(* IEC 61131-3 sources: podajnik-arkuszy/plc, 8 files *)

(* ---- FB_EStop.st ---- *)
(* Zezwolenie ruchu. Po otwarciu obwodu bezpieczenstwa i po wlaczeniu zasilania
   wymagane jest zbocze kasowania. Sam powrot styku bezpieczenstwa nie uruchamia maszyny. *)
FUNCTION_BLOCK FB_EStop
VAR_INPUT
    EStopOk : BOOL;
    Reset : BOOL;
END_VAR
VAR_OUTPUT
    RunEnable : BOOL;
END_VAR
VAR
    NeedReset : BOOL := TRUE;
END_VAR

IF NOT EStopOk THEN
    NeedReset := TRUE;
    RunEnable := FALSE;
ELSIF NeedReset THEN
    RunEnable := FALSE;
    IF Reset THEN
        NeedReset := FALSE;
        RunEnable := TRUE;
    END_IF;
ELSE
    RunEnable := TRUE;
END_IF;

END_FUNCTION_BLOCK

(* ---- FB_FuserBuckle.st ---- *)
(* Predkosc silnika fusera od czujnika wybrzuszenia przed nipem.
   Za duze wybrzuszenie: przyspiesz, zeby nie zgniesc arkusza.
   Za male: zwolnij, zeby nie rozmazac toneru na pasie.
   Waskie medium obcina predkosc. Zawiniecie na pasie zatrzymuje naped. *)
FUNCTION_BLOCK FB_FuserBuckle
VAR_INPUT
    Enable : BOOL;
    Nip : BOOL;
    BuckleHigh : BOOL;
    BuckleLow : BOOL;
    NarrowMedia : BOOL;
    Wrap : BOOL;
END_VAR
VAR_OUTPUT
    SpeedPct : INT;
    HeaterOn : BOOL;
    Jam : BOOL;
END_VAR

IF NOT Enable OR Wrap THEN
    SpeedPct := 0;
    HeaterOn := FALSE;
    Jam := Wrap;
ELSE
    Jam := FALSE;
    HeaterOn := TRUE; (* ceramika w pasie *)
    SpeedPct := 100;

    IF Nip AND BuckleHigh THEN
        SpeedPct := 130;
    ELSIF Nip AND BuckleLow THEN
        SpeedPct := 70;
    END_IF;

    IF NarrowMedia AND (SpeedPct > 80) THEN
        SpeedPct := 80;
    END_IF;
END_IF;

END_FUNCTION_BLOCK

(* ---- FB_FuserLife.st ---- *)
(* Licznik fusera. W XC4140 komplet type 01 (41X0253) wymienia sie po 150 000 stron.
   Ostrzezenie od 140 000. Kasowanie jest osobne od resetu zaciecia.
   Na panel idzie liczba tysiecy: rejestr 16-bit nie zmiesci 150000. *)
FUNCTION_BLOCK FB_FuserLife
VAR_INPUT
    SheetCount : INT;
    ResetService : BOOL;
END_VAR
VAR_OUTPUT
    Thousands : INT;
    Warn : BOOL;
    Due : BOOL;
END_VAR
VAR
    Total : DINT := 0;
    Prev : INT := 0;
    Seen : BOOL := FALSE;
END_VAR

IF NOT Seen THEN
    Prev := SheetCount;
    Seen := TRUE;
END_IF;

IF ResetService THEN
    Total := 0;
ELSIF SheetCount <> Prev THEN
    Total := Total + 1;
END_IF;
Prev := SheetCount;

IF Total > 150000 THEN
    Total := 150000;
END_IF;

Thousands := DINT_TO_INT(Total / 1000);
Warn := Total >= 140000;
Due := Total >= 150000;

END_FUNCTION_BLOCK

(* ---- FB_Motor.st ---- *)
(* Stycznik silnika. FaultIn przychodzi z termika.
   Gdy UseFeedback = TRUE, brak styku pomocniczego dluzej niz 500 ms jest awaria napedu. *)
FUNCTION_BLOCK FB_Motor
VAR_INPUT
    RunCmd : BOOL;
    Feedback : BOOL;
    UseFeedback : BOOL;
    FaultIn : BOOL;
    Reset : BOOL;
END_VAR
VAR_OUTPUT
    Run : BOOL;
    Fault : BOOL;
END_VAR
VAR
    TonFb : TON;
END_VAR

IF FaultIn THEN
    Fault := TRUE;
END_IF;

IF Reset AND NOT FaultIn THEN
    Fault := FALSE;
END_IF;

IF Fault THEN
    Run := FALSE;
    TonFb(IN := FALSE, PT := T#500ms);
ELSE
    IF UseFeedback THEN
        TonFb(IN := RunCmd AND NOT Feedback, PT := T#500ms);
    ELSE
        TonFb(IN := FALSE, PT := T#500ms);
    END_IF;

    IF TonFb.Q THEN
        Fault := TRUE;
        Run := FALSE;
    ELSE
        Run := RunCmd;
    END_IF;
END_IF;

END_FUNCTION_BLOCK

(* ---- FB_PID.st ---- *)
(* Regulator grzalki 24 V. Wyjscie 0..100 procent.
   Pierwszy cykl po wlaczeniu nie daje kopa od czlonu D. *)
FUNCTION_BLOCK FB_PID
VAR_INPUT
    Enable : BOOL;
    Setpoint : REAL;
    Actual : REAL;
    Kp : REAL;
    Ki : REAL;
    Kd : REAL;
    OutMin : REAL;
    OutMax : REAL;
    Cycle : REAL; (* okres obiegu w sekundach, przy cyklu 10 ms wpisz 0.01 *)
END_VAR
VAR_OUTPUT
    Out : REAL;
END_VAR
VAR
    Integral : REAL := 0.0;
    PrevError : REAL := 0.0;
    Armed : BOOL := FALSE;
    Error : REAL;
    Deriv : REAL;
    Raw : REAL;
END_VAR

IF NOT Enable OR (Cycle <= 0.0) THEN
    Integral := 0.0;
    PrevError := 0.0;
    Armed := FALSE;
    Out := 0.0;
ELSE
    Error := Setpoint - Actual;
    IF NOT Armed THEN
        PrevError := Error;
        Integral := 0.0;
        Armed := TRUE;
    END_IF;

    Integral := Integral + (Error * Cycle);
    Deriv := (Error - PrevError) / Cycle;
    PrevError := Error;
    Raw := (Kp * Error) + (Ki * Integral) + (Kd * Deriv);

    IF Raw > OutMax THEN
        Raw := OutMax;
        Integral := Integral - (Error * Cycle);
    ELSIF Raw < OutMin THEN
        Raw := OutMin;
        Integral := Integral - (Error * Cycle);
    END_IF;

    Out := Raw;
END_IF;

END_FUNCTION_BLOCK

(* ---- FB_SheetTrack.st ---- *)
(* Sciezka arkusza: sprzeglo podaje, czujnik wejscia, rejestracja, czujnik wyjscia.
   Brak czujnika w czasie JamTime (domyslnie 800 ms) = zaciecie.
   Przerwanie cyklu, gdy arkusz jest jeszcze na czujniku, tez jest zacieciem.
   Kasowanie dziala tylko przy pustej sciezce. *)
FUNCTION_BLOCK FB_SheetTrack
VAR_INPUT
    FeedCmd : BOOL;
    SensEntry : BOOL;
    SensRegister : BOOL;
    SensExit : BOOL;
    Reset : BOOL;
    JamTime : TIME := T#800ms;
END_VAR
VAR_OUTPUT
    MotorCmd : BOOL;
    Clutch : BOOL;
    AtRegister : BOOL;
    Jam : BOOL;
    Busy : BOOL;
    SheetCount : INT;
    PhaseOut : INT;
END_VAR
VAR
    Phase : INT := 0; (* 0 postoj, 1 czekam na rejestracje, 2 przejazd, 3 zejscie z czujnika *)
    TonReg : TON;
    TonExit : TON;
    rEntry : R_TRIG;
    rExit : R_TRIG;
END_VAR

rEntry(CLK := SensEntry);
rExit(CLK := SensExit);
TonReg(IN := (Phase = 1) AND NOT Jam, PT := JamTime);
TonExit(IN := (Phase = 2) AND NOT Jam, PT := JamTime);

IF Reset AND NOT SensEntry AND NOT SensRegister AND NOT SensExit THEN
    Jam := FALSE;
    Phase := 0;
END_IF;

IF Jam THEN
    MotorCmd := FALSE;
    Clutch := FALSE;
    AtRegister := FALSE;
ELSIF NOT FeedCmd AND (Phase <> 0) THEN
    IF SensEntry OR SensRegister OR SensExit THEN
        Jam := TRUE;
    ELSE
        Phase := 0;
    END_IF;
    MotorCmd := FALSE;
    Clutch := FALSE;
    AtRegister := FALSE;
ELSIF Phase = 0 THEN
    AtRegister := FALSE;
    IF FeedCmd AND rEntry.Q THEN
        Clutch := FALSE;
        MotorCmd := TRUE;
        Phase := 1;
    ELSIF FeedCmd AND (SensEntry OR SensRegister OR SensExit) THEN
        Jam := TRUE;
        Clutch := FALSE;
        MotorCmd := FALSE;
    ELSIF FeedCmd THEN
        Clutch := TRUE;
        MotorCmd := TRUE;
    ELSE
        Clutch := FALSE;
        MotorCmd := FALSE;
    END_IF;
ELSIF Phase = 1 THEN
    Clutch := FALSE;
    MotorCmd := TRUE;
    AtRegister := FALSE;
    IF SensRegister THEN
        Phase := 2;
        AtRegister := TRUE;
    ELSIF TonReg.Q THEN
        Jam := TRUE;
        Phase := 0;
        MotorCmd := FALSE;
    END_IF;
ELSIF Phase = 2 THEN
    Clutch := FALSE;
    MotorCmd := TRUE;
    AtRegister := TRUE;
    IF rExit.Q THEN
        SheetCount := SheetCount + 1;
        Phase := 3;
        AtRegister := FALSE;
    ELSIF TonExit.Q THEN
        Jam := TRUE;
        Phase := 0;
        MotorCmd := FALSE;
        AtRegister := FALSE;
    END_IF;
ELSE
    Clutch := FALSE;
    AtRegister := FALSE;
    MotorCmd := TRUE;
    IF NOT SensExit AND NOT SensEntry AND NOT SensRegister THEN
        Phase := 0;
        MotorCmd := FALSE;
    END_IF;
END_IF;

IF Jam THEN
    MotorCmd := FALSE;
    Clutch := FALSE;
    AtRegister := FALSE;
END_IF;

Busy := Jam OR (Phase <> 0) OR Clutch;
PhaseOut := Phase;

END_FUNCTION_BLOCK

(* ---- FB_Warmup.st ---- *)
(* Zezwolenie na podanie, gdy rolka 24 V jest w pasmie.
   Zadanie regulatora to 80 C. Ponizej 70 C start jest martwy.
   Powyzej 95 C to przegrzanie: grzalka odpada, nowy arkusz tez. *)
FUNCTION_BLOCK FB_Warmup
VAR_INPUT
    Enable : BOOL;
    Actual : REAL;
END_VAR
VAR_OUTPUT
    Ready : BOOL;
    Heating : BOOL;
    Overtemp : BOOL;
END_VAR

Overtemp := Enable AND (Actual > 95.0);
Ready := Enable AND (Actual >= 70.0) AND (Actual <= 95.0);
Heating := Enable AND (Actual < 70.0);

END_FUNCTION_BLOCK

(* ---- MAIN.st ---- *)
(* Podajnik arkuszy.
   OpenPLC Editor albo CODESYS: wklej FB_*.st jako bloki funkcyjne, a ten plik jako program.
   Cykl zadania: 10 ms.
   Adresy sa zgodne z electrical/io_map.csv.
   UseFeedback ustaw na TRUE dopiero po podpieciu styku pomocniczego stycznika pod I_MotorAux. *)
PROGRAM Main
VAR
    I_EstopOk AT %IX0.0 : BOOL;
    I_CoverClosed AT %IX0.1 : BOOL;
    I_SensEntry AT %IX0.2 : BOOL;
    I_SensRegister AT %IX0.3 : BOOL;
    I_SensExit AT %IX0.4 : BOOL;
    I_MotorFault AT %IX0.5 : BOOL;
    I_Start AT %IX0.6 : BOOL;
    I_Stop AT %IX0.7 : BOOL;
    I_Reset AT %IX1.0 : BOOL;
    I_MotorAux AT %IX1.1 : BOOL;
    I_FuserReset AT %IX1.2 : BOOL;
    I_Nip AT %IX1.3 : BOOL;
    I_BuckleHigh AT %IX1.4 : BOOL;
    I_BuckleLow AT %IX1.5 : BOOL;
    I_NarrowMedia AT %IX1.6 : BOOL;
    I_FuserWrap AT %IX1.7 : BOOL;
    IW_TempRaw AT %IW2 : INT;

    Q_Motor AT %QX0.0 : BOOL;
    Q_Clutch AT %QX0.1 : BOOL;
    Q_Gate AT %QX0.2 : BOOL;
    Q_LampRun AT %QX0.3 : BOOL;
    Q_LampFault AT %QX0.4 : BOOL;
    Q_Heater AT %QX0.5 : BOOL;
    Q_FuserMotor AT %QX0.6 : BOOL;

    QW_Heater AT %QW0 : INT; (* 0..1000 = 0.0..100.0 % *)
    QW_State AT %QW1 : INT;
    QW_Sheets AT %QW2 : INT;
    QW_Temp AT %QW3 : INT;
    QW_FuserK AT %QW4 : INT; (* tysiace stron od resetu fusera *)
    QW_FuserSvc AT %QW5 : INT; (* 0 ok, 1 ostrzezenie, 2 wymiana *)
    QW_FuserSpeed AT %QW6 : INT; (* procent predkosci silnika fusera *)
    QW_Warm AT %QW7 : INT; (* 0 zimna, 1 gotowa, 2 przegrzanie *)

    EStop : FB_EStop;
    Drive : FB_Motor;
    Track : FB_SheetTrack;
    Heat : FB_PID;
    FuserLife : FB_FuserLife;
    Buckle : FB_FuserBuckle;
    Warmup : FB_Warmup;
    rStart : R_TRIG;
    rStop : R_TRIG;
    rReset : R_TRIG;
    RunRequest : BOOL := FALSE;
    UseFeedback : BOOL := FALSE;
    MotionOk : BOOL;
    TempC : REAL;
    State : INT;
END_VAR

rStart(CLK := I_Start);
rStop(CLK := I_Stop);
rReset(CLK := I_Reset);

EStop(EStopOk := I_EstopOk, Reset := rReset.Q);

IF rStop.Q OR (NOT EStop.RunEnable) OR I_MotorFault OR (NOT I_CoverClosed) THEN
    RunRequest := FALSE;
END_IF;

MotionOk := EStop.RunEnable AND I_CoverClosed AND NOT I_MotorFault AND NOT Track.Jam;

FuserLife(SheetCount := Track.SheetCount, ResetService := I_FuserReset);
Buckle(
    Enable := EStop.RunEnable AND I_CoverClosed AND NOT FuserLife.Due,
    Nip := I_Nip,
    BuckleHigh := I_BuckleHigh,
    BuckleLow := I_BuckleLow,
    NarrowMedia := I_NarrowMedia,
    Wrap := I_FuserWrap
);

TempC := INT_TO_REAL(IW_TempRaw) / 10.0;
Warmup(
    Enable := EStop.RunEnable AND I_CoverClosed AND NOT FuserLife.Due,
    Actual := TempC
);

IF Warmup.Overtemp THEN
    RunRequest := FALSE;
END_IF;

IF rStart.Q AND MotionOk AND NOT Track.Busy AND NOT FuserLife.Due AND NOT Buckle.Jam AND Warmup.Ready THEN
    RunRequest := TRUE;
END_IF;

Track(
    FeedCmd := RunRequest AND MotionOk,
    SensEntry := I_SensEntry,
    SensRegister := I_SensRegister,
    SensExit := I_SensExit,
    Reset := rReset.Q,
    JamTime := T#800ms
);

Drive(
    RunCmd := Track.MotorCmd AND MotionOk,
    Feedback := I_MotorAux,
    UseFeedback := UseFeedback,
    FaultIn := I_MotorFault,
    Reset := rReset.Q
);

Heat(
    Enable := EStop.RunEnable AND I_CoverClosed AND NOT Track.Jam AND NOT Drive.Fault AND NOT Warmup.Overtemp,
    Setpoint := 80.0,
    Actual := TempC,
    Kp := 4.0,
    Ki := 0.8,
    Kd := 0.1,
    OutMin := 0.0,
    OutMax := 100.0,
    Cycle := 0.01
);

IF NOT EStop.RunEnable THEN
    State := 7;
ELSIF Drive.Fault OR I_MotorFault OR Warmup.Overtemp THEN
    State := 6;
ELSIF Buckle.Jam OR Track.Jam THEN
    State := 5;
ELSIF NOT I_CoverClosed THEN
    State := 8;
ELSIF Track.PhaseOut = 1 THEN
    State := 3;
ELSIF (Track.PhaseOut = 2) OR (Track.PhaseOut = 3) THEN
    State := 4;
ELSIF Track.Clutch THEN
    State := 2;
ELSE
    State := 1;
END_IF;

Q_Motor := Drive.Run AND EStop.RunEnable;
Q_Clutch := Track.Clutch AND EStop.RunEnable AND I_CoverClosed AND NOT Track.Jam;
Q_Gate := Track.AtRegister AND EStop.RunEnable AND I_CoverClosed AND NOT Track.Jam;
Q_LampRun := Q_Motor;
Q_LampFault := Track.Jam OR Drive.Fault OR NOT EStop.RunEnable OR FuserLife.Due OR Buckle.Jam OR Warmup.Overtemp;
Q_Heater := (Heat.Out > 1.0) AND Buckle.HeaterOn;
Q_FuserMotor := Buckle.SpeedPct > 0;

QW_Heater := REAL_TO_INT(Heat.Out * 10.0);
QW_State := State;
QW_Sheets := Track.SheetCount;
QW_Temp := IW_TempRaw;
QW_FuserK := FuserLife.Thousands;
IF FuserLife.Due THEN
    QW_FuserSvc := 2;
ELSIF FuserLife.Warn THEN
    QW_FuserSvc := 1;
ELSE
    QW_FuserSvc := 0;
END_IF;
QW_FuserSpeed := Buckle.SpeedPct;
IF Warmup.Overtemp THEN
    QW_Warm := 2;
ELSIF Warmup.Ready THEN
    QW_Warm := 1;
ELSE
    QW_Warm := 0;
END_IF;

END_PROGRAM
